(* Logix 5000 project; controller lab7 vendor 1 type 14 code 149 rev 32.11; software revision 32.00 *)

TASK MainTask (continuous, watchdog 500 ms) : MainProgram

MODULES
   Local : vendor 1 type 14 code 149 (Compact 0, rev 32.11)
      Discrete_IO : Embedded (Compact 1, rev 3.1, Output RPI 20 ms)
END_MODULES

PROGRAM MainProgram   (* main routine MainRoutine *)
VAR
   button_press : BOOL;
   conveyor_bit : BOOL;
   Green_button : ALIAS FOR Local:1:I.Data.2;
   left_green_light : ALIAS FOR Local:1:O.Data.2;
   ons : BOOL;
   red_button : ALIAS FOR Local:1:I.Data.1;
   red_light : ALIAS FOR Local:1:O.Data.0;
   right_green_light : ALIAS FOR Local:1:O.Data.5;
   system_run : BOOL;
   timer1 : TIMER := (PRE := 10000);
   timer2 : TIMER := (PRE := 500);
   timer3 : TIMER := (PRE := 500);
END_VAR

ROUTINE MainRoutine   (* ladder *)
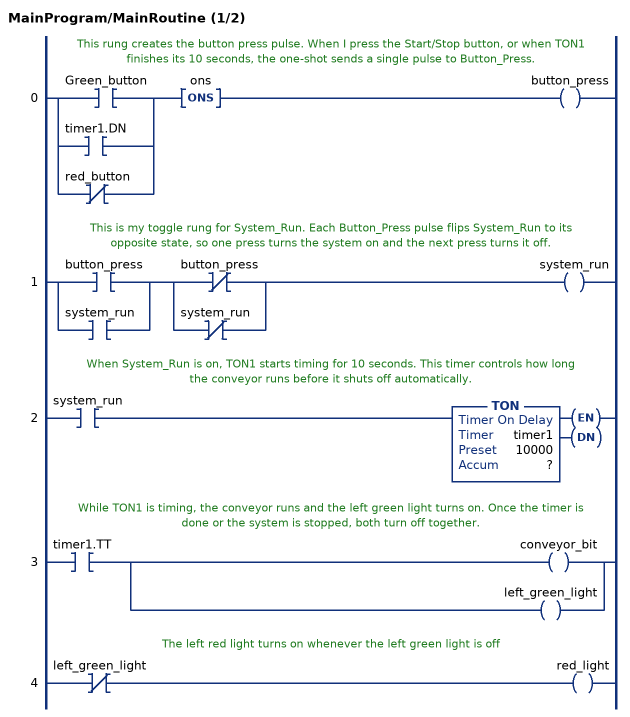
   // This rung creates the button press pulse. When I press the Start/Stop button, or when TON1 finishes its 10 seconds, the one-shot sends a single pulse to Button_Press.
   0: [XIC(Green_button) ,[XIC(timer1.DN) ,XIO(red_button) ] ]ONS(ons)OTE(button_press);
   // This is my toggle rung for System_Run. Each Button_Press pulse flips System_Run to its opposite state, so one press turns the system on and the next press turns it off.
   1: [XIC(button_press) ,XIC(system_run) ][XIO(button_press) ,XIO(system_run) ]OTE(system_run);
   // When System_Run is on, TON1 starts timing for 10 seconds. This timer controls how long the conveyor runs before it shuts off automatically.
   2: XIC(system_run)TON(timer1,?,?);
   // While TON1 is timing, the conveyor runs and the left green light turns on. Once the timer is done or the system is stopped, both turn off together.
   3: XIC(timer1.TT)[OTE(conveyor_bit) ,OTE(left_green_light) ];
   // The left red light turns on whenever the left green light is off
   4: XIO(left_green_light)OTE(red_light);
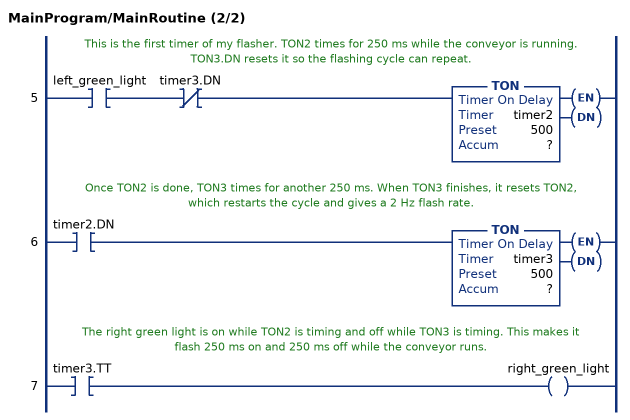
   // This is the first timer of my flasher. TON2 times for 250 ms while the conveyor is running. TON3.DN resets it so the flashing cycle can repeat.
   5: XIC(left_green_light)XIO(timer3.DN)TON(timer2,?,?);
   // Once TON2 is done, TON3 times for another 250 ms. When TON3 finishes, it resets TON2, which restarts the cycle and gives a 2 Hz flash rate.
   6: XIC(timer2.DN)TON(timer3,?,?);
   // The right green light is on while TON2 is timing and off while TON3 is timing. This makes it flash 250 ms on and 250 ms off while the conveyor runs.
   7: XIC(timer3.TT)OTE(right_green_light);
END_ROUTINE
END_PROGRAM
